Fanuc KAREL source: ka00122.KL

-- PROVISIONAL review KL for V940-1; original PC SHA256 7ee1c5de5b39a82df4ed0baa52f68e7e98ed9806811775d38306e1435918fcf7
-- Incomplete behavior may be omitted. Consult companion uncertainty JSON. Do not deploy.
PROGRAM KA00122
%NOLOCKGROUP
VAR
  DST : REAL
-- UNRESOLVED_DECL SRC type=002018
BEGIN
  -- V9_ZERO_TABLE_METADATA_HINT layout=0001; no indexed target words; source/name/runtime held
  -- UNRESOLVED_PC offsets 5-19; opcodes 2E,22,9D,33,B2
  -- UNRESOLVED_PC offsets 24-40; opcodes 22,9D,33,B1,64,23
  -- UNRESOLVED_PC offsets 45-49; opcodes 7F
END KA00122
